Fanuc KAREL source: KT00489.KL

PROGRAM KT00489
%NOLOCKGROUP
VAR
  P1: POSITION
  P2: JOINTPOS
  OUT: POSITION
BEGIN
  OUT = P1 : P2
END KT00489
